SUBAPPLICATION Uebung_094c2_AX (* Wie Uebung_094c_AX, aber mit MyLib::sys::NumericValue_TO_AUI2 als wiederverwendbarem Baustein statt der 2x inline duplizierten Kette (NumericValue_IDA+AD_TO_AUI+AUI_TO_AUI2+AUI_TO_AUDI+Q_NumericValue_AUDI je Dropdown). *)
  (* Standard: 61499-2; Description: Copyright (c) 2026 Meisterschulen am Ostbahnhof This program and the accompanying materials are made available under the terms of the Eclipse Public License 2.0 which is available at https://www.eclipse.org/legal/epl-2.0/ SPDX-License-Identifier: EPL-2.0 *)
  (* Version 1.0, 2026-10-13, Franz Höpfinger, Meisterschulen am Ostbahnhof, 2. Version von Uebung_094c_AX: die pro Dropdown duplizierte Lese/Echo-Kette wurde nach MyLib::sys::NumericValue_TO_AUI2 ausgelagert (u16ObjId als SubApp-Parameter statt fest verdrahtet). *)
  PACKAGE Uebungen;
  IMPORT Uebungen::const::UT::DefaultPool::InputNumber_I1;
  IMPORT Uebungen::const::UT::DefaultPool::InputNumber_I2;
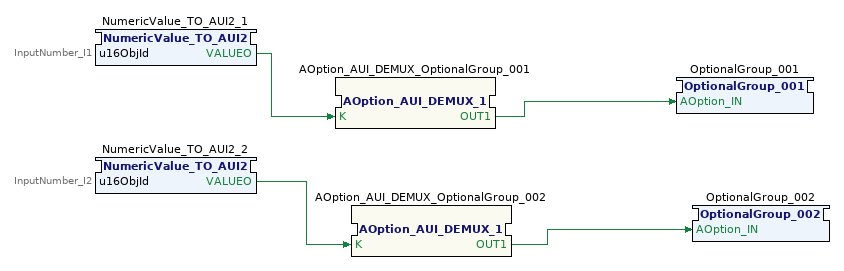
  FBS
    AOption_AUI_DEMUX_OptionalGroup_001 : Option::selection::AOption_AUI_DEMUX_1;
    AOption_AUI_DEMUX_OptionalGroup_002 : Option::selection::AOption_AUI_DEMUX_1;
  END_FBS
  SUBAPPS
    NumericValue_TO_AUI2_1 : MyLib::sys::NumericValue_TO_AUI2(u16ObjId := InputNumber_I1);
    NumericValue_TO_AUI2_2 : MyLib::sys::NumericValue_TO_AUI2(u16ObjId := InputNumber_I2);
    OptionalGroup_001 : MyLib_AX_Option::sys::OptionalGroup_001;
    OptionalGroup_002 : MyLib_AX_Option::sys::OptionalGroup_002;
  END_SUBAPPS
  ADAPTER_CONNECTIONS
    NumericValue_TO_AUI2_1.VALUEO TO AOption_AUI_DEMUX_OptionalGroup_001.K;
    NumericValue_TO_AUI2_2.VALUEO TO AOption_AUI_DEMUX_OptionalGroup_002.K;
    AOption_AUI_DEMUX_OptionalGroup_001.OUT1 TO OptionalGroup_001.AOption_IN;
    AOption_AUI_DEMUX_OptionalGroup_002.OUT1 TO OptionalGroup_002.AOption_IN;
  END_CONNECTIONS
END_SUBAPPLICATION
